(*
SPDX-FileCopyrightText: © 2026 Oleksandr Tiutyk <trofimich@gmail.com>
SPDX-License-Identifier: MIT
License: https://opensource.org/license/mit
*)

(*!
<summary>Binds external PLC variables to a freshly loaded workflow tree.</summary>
<description>
Invoked after the full tree is loaded, before variable requirement validation.
Must only modify variable bindings on the supplied fresh workflow.
</description>
*)
INTERFACE IWorkflowVariableBinder

(*!
<summary>Registers external PLC variables on the complete fresh tree before operand validation.</summary>
<param name="workflow">Loaded workflow instance.</param>
*)
METHOD BindVariables
VAR_INPUT
	workflow : IWorkflow;
END_VAR
END_METHOD

END_INTERFACE

(* stored: Version 1.1.0.1
   Itf IWorkflowVariableBinder: Id {940a7e41-3163-4c1d-9490-c9018d5b8999}
   Method BindVariables: Id {d3a0806a-146b-49fc-b0a7-37b7bdf2a1c2} *)
